// TIA Portal V21 export
// export: Created 2026-08-21T20:18:54.7477273Z, ExportSetting None, DisplayName Totally Integrated Automation Portal, DisplayVersion V21, DisplayName STEP 7 Professional, DisplayVersion V21, DisplayName STEP 7 Safety, DisplayVersion V21, DisplayName Tech WebApplication, DisplayVersion V21, DisplayName WinCC Basic/Comfort/Advanced, DisplayVersion V21, DisplayName WinCC Professional, DisplayVersion V21, DisplayName WinCC Unified, DisplayVersion V21
TYPE "UDT_MTP_BinProcessValueIn"
   STRUCT
      WQC { ExternalWritable := 'False'} : Byte := 16#FF;   // Worst Quality Code CCC
      V : Bool := false;   // External Source Value / Value
      VQC : Byte := 16#FF;   // Quality Code of the current received value
      VState0 { ExternalWritable := 'False'} : String[16] := '';   // Text Replacement Value (False) / text replacement for false
      VState1 { ExternalWritable := 'False'} : String[16] := '';   // Text Replacement Value (True) / text replacement for true
   END_STRUCT;
END_TYPE
